GLOBALCONSTANTS DefaultPool (* Global constants *)
  PACKAGE Uebungen::const::UT::Dialog;
  VAR_GLOBAL CONSTANT
    ISO_DESIGNATOR_WIDTH : UINT := 80;
    ISO_DESIGNATOR_HEIGHT : UINT := 80;
    ISO_MASK_SIZE : UINT := 480;
    ISO_VERSION_LABEL : STRING;
    MASK_WIDTH : UINT := 480;
    MASK_HEIGHT : UINT := 480;
    WorkingSet : UINT := 0;
    Macro_DataMask_M1 : UINT := 1;
    Macro_DataMask_M2 : UINT := 2;
    DataMask_M1 : UINT := 1000;
    DataMask_M2 : UINT := 1001;
    DataMask_Dlg_Vorlagen_invisible : UINT := 1002;
    Container_Dialog : UINT := 3400;
    Container_Dlg_Box : UINT := 3401;
    Container_Dlg_Icon_Info : UINT := 3402;
    Container_Dlg_Icon_Question : UINT := 3403;
    Container_Dlg_Icon_Warning : UINT := 3404;
    Container_Dlg_Icon_Error : UINT := 3405;
    Container_Dlg_Buttons_OK : UINT := 3410;
    Container_Dlg_Buttons_OKCancel : UINT := 3411;
    Container_Dlg_Buttons_AbortRetryIgnore : UINT := 3412;
    Container_Dlg_Buttons_YesNoCancel : UINT := 3413;
    Container_Dlg_Buttons_YesNo : UINT := 3414;
    Container_Dlg_Buttons_RetryCancel : UINT := 3415;
    SoftKeyMask_S1 : UINT := 4000;
    SoftKey_F1 : UINT := 5000;
    SoftKey_F2 : UINT := 5001;
    SoftKey_F3 : UINT := 5002;
    SoftKey_F4 : UINT := 5003;
    SoftKey_F5 : UINT := 5004;
    SoftKey_F6 : UINT := 5005;
    Button_Test1 : UINT := 6000;
    Button_Test2 : UINT := 6001;
    Button_Test3 : UINT := 6002;
    Button_Dlg_OK : UINT := 6900;
    Button_Dlg_Cancel : UINT := 6901;
    Button_Dlg_Abort : UINT := 6902;
    Button_Dlg_Retry : UINT := 6903;
    Button_Dlg_Ignore : UINT := 6904;
    Button_Dlg_Yes : UINT := 6905;
    Button_Dlg_No : UINT := 6906;
    OutputString_WorkingSet_0 : UINT := 11000;
    OutputString_SoftKey_F1 : UINT := 11001;
    OutputString_DataMask_M1 : UINT := 11013;
    OutputString_Result : UINT := 11014;
    OutputString_DataMask_M2 : UINT := 11015;
    OutputString_Button_Test1 : UINT := 11016;
    OutputString_Button_Test2 : UINT := 11017;
    OutputString_Button_Test3 : UINT := 11018;
    OutputString_Text_Toast : UINT := 11020;
    OutputString_Text_OK : UINT := 11021;
    OutputString_Text_Frage : UINT := 11022;
    OutputString_Dlg_Btn_OK : UINT := 11400;
    OutputString_Dlg_Btn_Cancel : UINT := 11401;
    OutputString_Dlg_Btn_Abort : UINT := 11402;
    OutputString_Dlg_Btn_Retry : UINT := 11403;
    OutputString_Dlg_Btn_Ignore : UINT := 11404;
    OutputString_Dlg_Btn_Yes : UINT := 11405;
    OutputString_Dlg_Btn_No : UINT := 11406;
    OutputString_Dlg_Title_Info : UINT := 11410;
    OutputString_Dlg_Title_Question : UINT := 11411;
    OutputString_Dlg_Title_Warning : UINT := 11412;
    OutputString_Dlg_Title_Error : UINT := 11413;
    OutputString_Dlg_Icon_Info : UINT := 11420;
    OutputString_Dlg_Icon_Question : UINT := 11421;
    OutputString_Dlg_Icon_Warning : UINT := 11422;
    OutputString_Dlg_Icon_Error : UINT := 11423;
    OutputString_SoftKey_F2 : UINT := 11501;
    OutputString_SoftKey_F3 : UINT := 11502;
    OutputString_SoftKey_F4 : UINT := 11503;
    OutputString_SoftKey_F5 : UINT := 11504;
    OutputString_SoftKey_F6 : UINT := 11505;
    OutputNumber_Result : UINT := 12000;
    Rectangle_Dlg_Cover : UINT := 14400;
    Rectangle_Dlg_Shadow : UINT := 14401;
    Rectangle_Dlg_Background : UINT := 14402;
    Rectangle_Dlg_Titlebar : UINT := 14403;
    Ellipse_Dlg_Icon_Info : UINT := 15400;
    Ellipse_Dlg_Icon_Question : UINT := 15401;
    Ellipse_Dlg_Icon_Warning : UINT := 15402;
    Ellipse_Dlg_Icon_Error : UINT := 15403;
    Logos_icon : UINT := 20500;
    FontAttributes_6x8 : UINT := 23000;
    FontAttributes_8x12 : UINT := 23001;
    FontAttributes_Dlg_8x12_black : UINT := 23400;
    FontAttributes_Dlg_8x12_white : UINT := 23401;
    FontAttributes_Dlg_12x16_white : UINT := 23402;
    FontAttributes_Dlg_12x16_black : UINT := 23403;
    LineAttributes_Dlg_none_white : UINT := 24400;
    LineAttributes_Dlg_Frame : UINT := 24401;
    LineAttributes_Dlg_none_grey : UINT := 24402;
    FillAttributes_Dlg_White : UINT := 25400;
    FillAttributes_Dlg_Shadow : UINT := 25401;
    FillAttributes_Dlg_Title : UINT := 25402;
    FillAttributes_Dlg_Icon_Info : UINT := 25403;
    FillAttributes_Dlg_Icon_Question : UINT := 25404;
    FillAttributes_Dlg_Icon_Warning : UINT := 25405;
    FillAttributes_Dlg_Icon_Error : UINT := 25406;
    ObjectPointer_Dlg_Cover : UINT := 27900;
    ObjectPointer_Dlg_Icon : UINT := 27901;
    ObjectPointer_Dlg_Title : UINT := 27902;
    ObjectPointer_Dlg_Text : UINT := 27903;
    ObjectPointer_Dlg_Buttons : UINT := 27904;
    AuxFunction2_X1 : UINT := 31000;
  END_VAR
END_GLOBALCONSTANTS
